(* IEC 61131-3 sources: kns-port-domestic/targets/astra/src/POUs/Model/FB_StormGenerator, 11 files *)

(* ---- FB_StormGenerator.decl.st ---- *)
// Назначение: ливни модели по seed. На сутки d — начальное состояние x0 = udiSeed XOR (d · 16#9E3779B9),
//             равномерные u = (x AND 16#00FFFFFF) / 2^24 по шагам F_Xorshift32: число ливней
//             0…uiStormsPerDayMax, для каждого — начало (равномерно в сутках), длительность (между
//             tDurationMin и tDurationMax), пик (между rPeakMin_m3h и rPeakMax_m3h). Форма — трапеция:
//             рост 15 %, полка 50 %, спад 35 % длительности. Ливни зависят только от seed и номера
//             суток — одинаковы при любом ускорении и шаге вызова. Ливень предыдущих суток, который
//             не закончился к полуночи, продолжается. StartNow — внеочередной ливень той же формы,
//             Clear — снять идущие ливни (xResetPlant).
// Автор:      kr0nsch
// Версия:     0.1.0
// Документ:   docs/DESIGN.md, раздел 11.2
FUNCTION_BLOCK FB_StormGenerator
VAR_INPUT
    lrClock_h         : LREAL;      // часы модели: ч от полуночи суток 0
    udiSeed           : UDINT;      // stSimCfg.udiSeed
    uiStormsPerDayMax : UINT;       // не больше SIM_STORMS_MAX (больше — ограничивается)
    rPeakMin_m3h      : REAL;
    rPeakMax_m3h      : REAL;
    tDurationMin      : TIME;
    tDurationMax      : TIME;
END_VAR
VAR_OUTPUT
    rInflow_m3h : REAL;             // приток ливней сейчас
    xActive     : BOOL;             // идёт хотя бы один ливень
    udiDay      : UDINT;            // номер суток модели
    uiCount     : UINT;             // ливней в текущих сутках
    astStorm    : ARRAY[1..GVL_Const.SIM_STORMS_MAX] OF ST_StormEvent;   // ливни текущих суток, 1…uiCount
END_VAR
VAR
    astPrev     : ARRAY[1..GVL_Const.SIM_STORMS_MAX] OF ST_StormEvent;   // ливни предыдущих суток
    uiPrevCount : UINT;
    astWork     : ARRAY[1..GVL_Const.SIM_STORMS_MAX] OF ST_StormEvent;   // результат Generate
    dwState     : DWORD;            // состояние генератора при заполнении суток
    xGenerated  : BOOL;             // ливни заполнены для udiDayGen и параметров ниже
    udiDayGen   : UDINT;
    udiSeedGen  : UDINT;
    uiMaxGen    : UINT;
    rPeakMinGen : REAL;
    rPeakMaxGen : REAL;
    tMinGen     : TIME;
    tMaxGen     : TIME;
    xManual     : BOOL;             // внеочередной ливень (StartNow) ещё не закончился
    stManual    : ST_StormEvent;    // его длительность и пик
    lrManualStart_h : LREAL;        // его начало по часам модели
    lrSuppress_h : LREAL := -1.0;   // ливни, начавшиеся раньше этого момента, сняты (Clear)
    uiStorm     : UINT;             // индекс ливня
    lrStart_h   : LREAL;            // начало ливня по часам модели
END_VAR

(* ---- AddStorm.method.decl.st ---- *)
// Добавить к rInflow_m3h приток ливня (трапеция: рост 15 %, полка 50 %, спад 35 %) в момент lrClock_h;
// ливень идёт — xActive. Вне [начало, начало + длительность) ливень ничего не добавляет
METHOD PRIVATE AddStorm
VAR_INPUT
    lrStartAt_h : LREAL;    // начало ливня по часам модели
    tDur        : TIME;     // длительность
    rPeak       : REAL;     // пик, м³/ч
END_VAR
VAR
    lrTau_s  : LREAL;       // время от начала ливня
    lrDur_s  : LREAL;       // длительность, с
    lrRise_s : LREAL;       // конец роста
    lrFall_s : LREAL;       // начало спада
END_VAR

(* ---- AddStorm.method.impl.st ---- *)
lrDur_s := PL.F_TimeToSec(tIn := tDur);
lrTau_s := (lrClock_h - lrStartAt_h) * REAL_TO_LREAL(GVL_Const.SIM_S_PER_H);
IF lrDur_s <= 0.0 OR lrTau_s < 0.0 OR lrTau_s >= lrDur_s THEN
    RETURN;
END_IF

xActive := TRUE;
lrRise_s := REAL_TO_LREAL(GVL_Const.SIM_STORM_RISE_SHARE) * lrDur_s;
lrFall_s := (1.0 - REAL_TO_LREAL(GVL_Const.SIM_STORM_FALL_SHARE)) * lrDur_s;
IF lrTau_s < lrRise_s THEN
    rInflow_m3h := rInflow_m3h + LREAL_TO_REAL(REAL_TO_LREAL(rPeak) * lrTau_s / lrRise_s);
ELSIF lrTau_s < lrFall_s THEN
    rInflow_m3h := rInflow_m3h + rPeak;
ELSE
    rInflow_m3h := rInflow_m3h
                   + LREAL_TO_REAL(REAL_TO_LREAL(rPeak) * (lrDur_s - lrTau_s) / (lrDur_s - lrFall_s));
END_IF

(* ---- Clear.method.decl.st ---- *)
// Снять ливни (stSimCmd.xResetPlant): ливни, начавшиеся раньше lrFrom_h, и внеочередной ливень
// больше не дают притока; ливни генератора, которые начнутся позже, идут как обычно
METHOD PUBLIC Clear
VAR_INPUT
    lrFrom_h : LREAL;       // момент снятия по часам модели (обычно текущие часы)
END_VAR

(* ---- FB_StormGenerator.impl.st ---- *)
// 1. Сутки модели (часы не бывают отрицательными: модель начинает с 0…24 ч)
IF lrClock_h > 0.0 THEN
    udiDay := FloorU(lrValue := lrClock_h / REAL_TO_LREAL(GVL_Const.SIM_HOURS_PER_DAY));
ELSE
    udiDay := 0;
END_IF

// 2. Ливни текущих и предыдущих суток — заново при смене суток или параметров генератора
IF NOT xGenerated OR udiDay <> udiDayGen OR udiSeed <> udiSeedGen OR uiStormsPerDayMax <> uiMaxGen
   OR rPeakMin_m3h <> rPeakMinGen OR rPeakMax_m3h <> rPeakMaxGen OR tDurationMin <> tMinGen
   OR tDurationMax <> tMaxGen THEN
    uiCount := Generate(udiForDay := udiDay);
    astStorm := astWork;
    IF udiDay > 0 THEN
        uiPrevCount := Generate(udiForDay := udiDay - 1);
        astPrev := astWork;
    ELSE
        uiPrevCount := 0;
    END_IF
    xGenerated := TRUE;
    udiDayGen := udiDay;
    udiSeedGen := udiSeed;
    uiMaxGen := uiStormsPerDayMax;
    rPeakMinGen := rPeakMin_m3h;
    rPeakMaxGen := rPeakMax_m3h;
    tMinGen := tDurationMin;
    tMaxGen := tDurationMax;
END_IF

// 3. Приток: сумма трапеций идущих ливней; ливни, начавшиеся до Clear, сняты
rInflow_m3h := 0.0;
xActive := FALSE;
FOR uiStorm := 1 TO uiPrevCount DO
    lrStart_h := UDINT_TO_LREAL(udiDay - 1) * REAL_TO_LREAL(GVL_Const.SIM_HOURS_PER_DAY)
                 + REAL_TO_LREAL(astPrev[uiStorm].rStart_h);
    IF lrStart_h >= lrSuppress_h THEN
        AddStorm(lrStartAt_h := lrStart_h, tDur := astPrev[uiStorm].tDuration, rPeak := astPrev[uiStorm].rPeak_m3h);
    END_IF
END_FOR
FOR uiStorm := 1 TO uiCount DO
    lrStart_h := UDINT_TO_LREAL(udiDay) * REAL_TO_LREAL(GVL_Const.SIM_HOURS_PER_DAY)
                 + REAL_TO_LREAL(astStorm[uiStorm].rStart_h);
    IF lrStart_h >= lrSuppress_h THEN
        AddStorm(lrStartAt_h := lrStart_h, tDur := astStorm[uiStorm].tDuration, rPeak := astStorm[uiStorm].rPeak_m3h);
    END_IF
END_FOR
IF xManual THEN
    IF (lrClock_h - lrManualStart_h) * REAL_TO_LREAL(GVL_Const.SIM_S_PER_H)
       >= PL.F_TimeToSec(tIn := stManual.tDuration) THEN
        xManual := FALSE;       // внеочередной ливень закончился
    ELSE
        AddStorm(lrStartAt_h := lrManualStart_h, tDur := stManual.tDuration, rPeak := stManual.rPeak_m3h);
    END_IF
END_IF

(* ---- FloorU.method.decl.st ---- *)
// Целая часть неотрицательного LREAL (LREAL_TO_UDINT округляет — поправка вниз); отрицательное — 0
METHOD PRIVATE FloorU : UDINT
VAR_INPUT
    lrValue : LREAL;        // значение, ≥ 0
END_VAR
VAR
    udiRound : UDINT;       // округлённое значение
END_VAR

(* ---- FloorU.method.impl.st ---- *)
IF lrValue <= 0.0 THEN
    FloorU := 0;
    RETURN;
END_IF
udiRound := LREAL_TO_UDINT(lrValue);
IF UDINT_TO_LREAL(udiRound) > lrValue THEN
    udiRound := udiRound - 1;
END_IF
FloorU := udiRound;

(* ---- Generate.method.decl.st ---- *)
// Ливни суток udiForDay в astWork; результат — их число. Порядок выборок: число ливней, затем для
// каждого — начало, длительность, пик (так же в эталоне tools_project/plant_reference.py)
METHOD PRIVATE Generate : UINT
VAR_INPUT
    udiForDay : UDINT;      // номер суток
END_VAR
VAR
    uiMax    : UINT;        // предел числа ливней
    uiN      : UINT;        // число ливней
    uiK      : UINT;        // индекс ливня
    lrMin_ms : LREAL;       // границы длительности, мс
    lrMax_ms : LREAL;
    rLoPeak  : REAL;        // границы пика (упорядоченные)
    rHiPeak  : REAL;
END_VAR

(* ---- Generate.method.impl.st ---- *)
// начальное состояние суток; UDINT-умножение — по модулю 2^32
dwState := UDINT_TO_DWORD(udiSeed) XOR UDINT_TO_DWORD(udiForDay * GVL_Const.SIM_SEED_DAY_MUL);
IF dwState = 0 THEN
    dwState := GVL_Const.SIM_XS_ZERO_STATE;
END_IF

uiMax := MIN(uiStormsPerDayMax, GVL_Const.SIM_STORMS_MAX);
uiN := UDINT_TO_UINT(FloorU(lrValue := Draw() * UINT_TO_LREAL(uiMax + 1)));
uiN := MIN(uiN, uiMax);

lrMin_ms := UDINT_TO_LREAL(TIME_TO_UDINT(MIN(tDurationMin, tDurationMax)));
lrMax_ms := UDINT_TO_LREAL(TIME_TO_UDINT(MAX(tDurationMin, tDurationMax)));
rLoPeak := MIN(rPeakMin_m3h, rPeakMax_m3h);
rHiPeak := MAX(rPeakMin_m3h, rPeakMax_m3h);
FOR uiK := 1 TO uiN DO
    astWork[uiK].rStart_h := LREAL_TO_REAL(Draw() * REAL_TO_LREAL(GVL_Const.SIM_HOURS_PER_DAY));
    astWork[uiK].tDuration := UDINT_TO_TIME(LREAL_TO_UDINT(lrMin_ms + Draw() * (lrMax_ms - lrMin_ms)));
    astWork[uiK].rPeak_m3h := LREAL_TO_REAL(REAL_TO_LREAL(rLoPeak) + Draw() * REAL_TO_LREAL(rHiPeak - rLoPeak));
END_FOR
Generate := uiN;

(* ---- StartNow.method.decl.st ---- *)
// Внеочередной ливень (stSimCmd.xStormNow): трапеция с пиком rPeak_m3h и длительностью tDuration
// от момента lrStartAt_h; заменяет предыдущий внеочередной ливень. Длительность 0 или пик ≤ 0 — не начинается
METHOD PUBLIC StartNow
VAR_INPUT
    lrStartAt_h : LREAL;    // начало по часам модели (обычно текущие часы)
    rPeak_m3h   : REAL;     // пик притока
    tDuration   : TIME;     // длительность
END_VAR

(* ---- StartNow.method.impl.st ---- *)
IF tDuration > T#0S AND rPeak_m3h > 0.0 AND PL.F_IsFinite(rIn := rPeak_m3h) THEN
    xManual := TRUE;
    lrManualStart_h := lrStartAt_h;
    stManual.rStart_h := 0.0;
    stManual.tDuration := tDuration;
    stManual.rPeak_m3h := rPeak_m3h;
ELSE
    xManual := FALSE;
END_IF
